Fanuc KAREL source: KD00039.KL

PROGRAM KD00039
%NOLOCKGROUP
VAR
  I: INTEGER
  J: INTEGER
  B: BOOLEAN
  R: REAL
  S: STRING[80]
BEGIN
  CONDITION[1]:
  WHEN DIN[1] = ON DO
    SIGNAL EVENT[1]
  ENDCONDITION
END KD00039
